(* IEC 61131-3 sources: codesys-framework/txt/application/WeVe Core (library)/60 Event/DUT, 3 files *)

(* ---- SC_Event.dut.st ---- *)
TYPE SC_Event :
STRUCT
	udiEventId 			: UDINT;
	nSubMachine 		: USINT;
	nSubMachineId 		: USINT;
	eEventLevel 		: E_EventLevels;
	xResetable 			: BOOL;		// TRUE = blijft actief tot Reset(), ook als de conditie weg is
	sMessage 			: STRING(GVL_Logger.cMaxMessageLength) := '';	// placeholders %0..%9
END_STRUCT
END_TYPE

(* ---- SC_EventPayload.dut.st ---- *)
TYPE SC_EventPayload :
STRUCT
	asPayload 	: ARRAY[0..9] OF STRING := [10('')];
END_STRUCT
END_TYPE

(* ---- SC_EventState.dut.st ---- *)
TYPE SC_EventState :
STRUCT
	xWarningIsOn 	: BOOL;
	xAlarmIsOn 		: BOOL;
END_STRUCT
END_TYPE
